// TIA Portal V20 export
TYPE "Afag_Variablen_Positionen_Dreh"
   STRUCT
      Start_POS_Position : Array[0..15] of Bool;
      POS_OK_Position : Array[0..15] of Bool;
      Soll_Wert_in_Grad_Position : Array[0..15] of Real;
      Soll_Speed_in_Prozent_Position : Array[0..15] of Int;
      Positionstoleranz_Position : Array[0..15] of Real;
      Soll_Beschleunigung_in_Grad_s_Position : Array[0..15] of Int;
      A_Softw_ES_min_Grad : Real;
      A_Softw_ES_max_Grad : Real;
      A_Max_Speed_Grad_s : Int;
      A_Max_Beschleunigung_Grad_s : Int;
   END_STRUCT;
   // Soll_Speed_in_Prozent_Position[0..15] := 10;
   // Positionstoleranz_Position[0..15] := 0.5;
   // Soll_Beschleunigung_in_Grad_s_Position[0..15] := 1450;
END_TYPE
